(* IEC 61131-3 sources: virtual-bottling-plant/plc/src/generated/bridge, 13 files *)

(* ---- Bridge_Alarms.st ---- *)
(* GENERATED by plc/scripts/gen_plc_io.py from contracts/modbus/plc-io.yaml. Do not edit by hand. *)
(* Alarm table: bit0 active, bit1 acked, bit2 first-out, bits 8-11 prio. *)
PROGRAM Bridge_Alarms
  VAR_EXTERNAL
    G_Alarms : ST_AlarmSummary;
  END_VAR
  VAR
    ALM_T101_BrixOutOfSpec AT %MW601 : INT;
    ALM_T101_CommsLost AT %MW602 : INT;
    ALM_P201_LowTemp AT %MW603 : INT;
    ALM_P201_SteamLow AT %MW604 : INT;
    ALM_P201_CommsLost AT %MW605 : INT;
    ALM_T301_LowLevel AT %MW606 : INT;
    ALM_T301_CommsLost AT %MW607 : INT;
    ALM_F401_NozzleLeak AT %MW608 : INT;
    ALM_F401_CommsLost AT %MW609 : INT;
    ALM_C501_Jam AT %MW610 : INT;
    ALM_C501_Breakdown AT %MW611 : INT;
    ALM_C501_CapsEmpty AT %MW612 : INT;
    ALM_C501_CommsLost AT %MW613 : INT;
    ALM_L601_RollEmpty AT %MW614 : INT;
    ALM_L601_LabelError AT %MW615 : INT;
    ALM_L601_Breakdown AT %MW616 : INT;
    ALM_L601_CommsLost AT %MW617 : INT;
    ALM_Q701_CommsLost AT %MW618 : INT;
    ALM_K801_Jam AT %MW619 : INT;
    ALM_K801_Breakdown AT %MW620 : INT;
    ALM_K801_CommsLost AT %MW621 : INT;
    ALM_LINE_CommsLost AT %MW622 : INT;
  END_VAR
  ALM_T101_BrixOutOfSpec := UINT_TO_INT(G_Alarms.W1);
  ALM_T101_CommsLost := UINT_TO_INT(G_Alarms.W2);
  ALM_P201_LowTemp := UINT_TO_INT(G_Alarms.W3);
  ALM_P201_SteamLow := UINT_TO_INT(G_Alarms.W4);
  ALM_P201_CommsLost := UINT_TO_INT(G_Alarms.W5);
  ALM_T301_LowLevel := UINT_TO_INT(G_Alarms.W6);
  ALM_T301_CommsLost := UINT_TO_INT(G_Alarms.W7);
  ALM_F401_NozzleLeak := UINT_TO_INT(G_Alarms.W8);
  ALM_F401_CommsLost := UINT_TO_INT(G_Alarms.W9);
  ALM_C501_Jam := UINT_TO_INT(G_Alarms.W10);
  ALM_C501_Breakdown := UINT_TO_INT(G_Alarms.W11);
  ALM_C501_CapsEmpty := UINT_TO_INT(G_Alarms.W12);
  ALM_C501_CommsLost := UINT_TO_INT(G_Alarms.W13);
  ALM_L601_RollEmpty := UINT_TO_INT(G_Alarms.W14);
  ALM_L601_LabelError := UINT_TO_INT(G_Alarms.W15);
  ALM_L601_Breakdown := UINT_TO_INT(G_Alarms.W16);
  ALM_L601_CommsLost := UINT_TO_INT(G_Alarms.W17);
  ALM_Q701_CommsLost := UINT_TO_INT(G_Alarms.W18);
  ALM_K801_Jam := UINT_TO_INT(G_Alarms.W19);
  ALM_K801_Breakdown := UINT_TO_INT(G_Alarms.W20);
  ALM_K801_CommsLost := UINT_TO_INT(G_Alarms.W21);
  ALM_LINE_CommsLost := UINT_TO_INT(G_Alarms.W22);
END_PROGRAM

(* ---- Bridge_C501.st ---- *)
(* GENERATED by plc/scripts/gen_plc_io.py from contracts/modbus/plc-io.yaml. Do not edit by hand. *)
(* Status block C501 (%MW200…). *)
PROGRAM Bridge_C501
  VAR_EXTERNAL
    G_In : ST_SimInputs;
    G_Out : ST_SimOutputs;
    G_Status : ST_Status;
    G_Comms : ST_CommsStatus;
    G_Alarms : ST_AlarmSummary;
  END_VAR
  VAR
    C501_State AT %MW200 : INT;
    C501_Mode AT %MW201 : INT;
    C501_StopReason AT %MW202 : INT;
    C501_AlarmWord AT %MW203 : INT;
    C501_CommsOk AT %MW204 : INT;
    C501_Blocked AT %MW205 : INT;
    C501_Starved AT %MW206 : INT;
    C501_Running AT %MW207 : INT;
    C501_Speed AT %MW208 : INT;
    C501_SpeedSP AT %MW209 : INT;
    C501_Torque AT %MW210 : INT;
    C501_LT502_CapHopper AT %MW211 : INT;
  END_VAR
  C501_State := PackMLStateToInt(G_Status.C501.State);
  C501_Mode := PackMLModeToInt(G_Status.C501.Mode);
  C501_StopReason := G_Status.C501.StopReason;
  C501_AlarmWord := G_Alarms.C501_Word;
  C501_CommsOk := BOOL_TO_INT(G_Comms.C501);
  C501_Blocked := BOOL_TO_INT(G_Status.C501.Blocked);
  C501_Starved := BOOL_TO_INT(G_Status.C501.Starved);
  C501_Running := BOOL_TO_INT(G_In.C501_Running);
  C501_Speed := REAL_TO_INT(G_In.C501_Speed);
  C501_SpeedSP := REAL_TO_INT(G_Out.C501_SpeedSP);
  C501_Torque := REAL_TO_INT(G_In.C501_Torque * 100.0);
  C501_LT502_CapHopper := REAL_TO_INT(G_In.LT502_CapHopper * 10.0);
END_PROGRAM

(* ---- Bridge_Commands.st ---- *)
(* GENERATED by plc/scripts/gen_plc_io.py from contracts/modbus/plc-io.yaml. Do not edit by hand. *)
(* One-shot commands: valid in G_Cmd for the scan they arrive, then 0. *)
PROGRAM Bridge_Commands
  VAR_EXTERNAL
    G_Cmd : ST_Commands;
  END_VAR
  VAR
    F401_Cmd AT %MW803 : INT;
    C501_Cmd AT %MW804 : INT;
    L601_Cmd AT %MW805 : INT;
    Q701_Cmd AT %MW806 : INT;
    K801_Cmd AT %MW807 : INT;
    LINE_Cmd AT %MW808 : INT;
    F401_StopReason AT %MW813 : INT;
    C501_StopReason AT %MW814 : INT;
    L601_StopReason AT %MW815 : INT;
    Q701_StopReason AT %MW816 : INT;
    K801_StopReason AT %MW817 : INT;
    AlarmAck AT %MW820 : INT;
    P201_TempSP AT %MW821 : INT;
  END_VAR
  G_Cmd.F401_Cmd := IntToCommand(F401_Cmd);
  F401_Cmd := 0;
  G_Cmd.C501_Cmd := IntToCommand(C501_Cmd);
  C501_Cmd := 0;
  G_Cmd.L601_Cmd := IntToCommand(L601_Cmd);
  L601_Cmd := 0;
  G_Cmd.Q701_Cmd := IntToCommand(Q701_Cmd);
  Q701_Cmd := 0;
  G_Cmd.K801_Cmd := IntToCommand(K801_Cmd);
  K801_Cmd := 0;
  G_Cmd.LINE_Cmd := IntToCommand(LINE_Cmd);
  LINE_Cmd := 0;
  G_Cmd.F401_StopReason := F401_StopReason;
  F401_StopReason := 0;
  G_Cmd.C501_StopReason := C501_StopReason;
  C501_StopReason := 0;
  G_Cmd.L601_StopReason := L601_StopReason;
  L601_StopReason := 0;
  G_Cmd.Q701_StopReason := Q701_StopReason;
  Q701_StopReason := 0;
  G_Cmd.K801_StopReason := K801_StopReason;
  K801_StopReason := 0;
  G_Cmd.AlarmAck := AlarmAck;
  AlarmAck := 0;
  G_Cmd.P201_TempSP := INT_TO_REAL(P201_TempSP) / 10.0;
  P201_TempSP := 0;
END_PROGRAM

(* ---- Bridge_Counters.st ---- *)
(* GENERATED by plc/scripts/gen_plc_io.py from contracts/modbus/plc-io.yaml. Do not edit by hand. *)
(* 32-bit counters (%MD, high word first on Modbus). *)
PROGRAM Bridge_Counters
  VAR_EXTERNAL
    G_In : ST_SimInputs;
    G_Counters : ST_Counters;
  END_VAR
  VAR
    F401_Count AT %MD0 : DINT;
    C501_Count AT %MD1 : DINT;
    L601_Count AT %MD2 : DINT;
    Q701_Count AT %MD3 : DINT;
    Q701_RejectCount AT %MD4 : DINT;
    Q701_GoodCount AT %MD5 : DINT;
    K801_CaseCount AT %MD6 : DINT;
    T101_ConcLotNo AT %MD7 : DINT;
    SIM_TimeMs AT %MD8 : DINT;
  END_VAR
  F401_Count := UDINT_TO_DINT(G_In.F401_Count);
  C501_Count := UDINT_TO_DINT(G_In.C501_Count);
  L601_Count := UDINT_TO_DINT(G_In.L601_Count);
  Q701_Count := UDINT_TO_DINT(G_In.Q701_Count);
  Q701_RejectCount := UDINT_TO_DINT(G_In.Q701_RejectCount);
  Q701_GoodCount := UDINT_TO_DINT(G_Counters.Q701_GoodCount);
  K801_CaseCount := UDINT_TO_DINT(G_In.K801_CaseCount);
  T101_ConcLotNo := UDINT_TO_DINT(G_In.T101_ConcLotNo);
  SIM_TimeMs := UDINT_TO_DINT(G_In.SIM_TimeMs);
END_PROGRAM

(* ---- Bridge_F401.st ---- *)
(* GENERATED by plc/scripts/gen_plc_io.py from contracts/modbus/plc-io.yaml. Do not edit by hand. *)
(* Status block F401 (%MW150…). *)
PROGRAM Bridge_F401
  VAR_EXTERNAL
    G_In : ST_SimInputs;
    G_Out : ST_SimOutputs;
    G_Status : ST_Status;
    G_Comms : ST_CommsStatus;
    G_Alarms : ST_AlarmSummary;
  END_VAR
  VAR
    F401_State AT %MW150 : INT;
    F401_Mode AT %MW151 : INT;
    F401_StopReason AT %MW152 : INT;
    F401_AlarmWord AT %MW153 : INT;
    F401_CommsOk AT %MW154 : INT;
    F401_Blocked AT %MW155 : INT;
    F401_Starved AT %MW156 : INT;
    F401_Running AT %MW157 : INT;
    F401_Speed AT %MW158 : INT;
    F401_SpeedSP AT %MW159 : INT;
    F401_FillTargetG AT %MW160 : INT;
  END_VAR
  F401_State := PackMLStateToInt(G_Status.F401.State);
  F401_Mode := PackMLModeToInt(G_Status.F401.Mode);
  F401_StopReason := G_Status.F401.StopReason;
  F401_AlarmWord := G_Alarms.F401_Word;
  F401_CommsOk := BOOL_TO_INT(G_Comms.F401);
  F401_Blocked := BOOL_TO_INT(G_Status.F401.Blocked);
  F401_Starved := BOOL_TO_INT(G_Status.F401.Starved);
  F401_Running := BOOL_TO_INT(G_In.F401_Running);
  F401_Speed := REAL_TO_INT(G_In.F401_Speed);
  F401_SpeedSP := REAL_TO_INT(G_Out.F401_SpeedSP);
  F401_FillTargetG := REAL_TO_INT(G_Out.F401_FillTargetG * 10.0);
END_PROGRAM

(* ---- Bridge_K801.st ---- *)
(* GENERATED by plc/scripts/gen_plc_io.py from contracts/modbus/plc-io.yaml. Do not edit by hand. *)
(* Status block K801 (%MW350…). *)
PROGRAM Bridge_K801
  VAR_EXTERNAL
    G_In : ST_SimInputs;
    G_Out : ST_SimOutputs;
    G_Status : ST_Status;
    G_Comms : ST_CommsStatus;
    G_Alarms : ST_AlarmSummary;
  END_VAR
  VAR
    K801_State AT %MW350 : INT;
    K801_Mode AT %MW351 : INT;
    K801_StopReason AT %MW352 : INT;
    K801_AlarmWord AT %MW353 : INT;
    K801_CommsOk AT %MW354 : INT;
    K801_Blocked AT %MW355 : INT;
    K801_Starved AT %MW356 : INT;
    K801_Running AT %MW357 : INT;
    K801_Speed AT %MW358 : INT;
    K801_SpeedSP AT %MW359 : INT;
  END_VAR
  K801_State := PackMLStateToInt(G_Status.K801.State);
  K801_Mode := PackMLModeToInt(G_Status.K801.Mode);
  K801_StopReason := G_Status.K801.StopReason;
  K801_AlarmWord := G_Alarms.K801_Word;
  K801_CommsOk := BOOL_TO_INT(G_Comms.K801);
  K801_Blocked := BOOL_TO_INT(G_Status.K801.Blocked);
  K801_Starved := BOOL_TO_INT(G_Status.K801.Starved);
  K801_Running := BOOL_TO_INT(G_In.K801_Running);
  K801_Speed := REAL_TO_INT(G_In.K801_Speed);
  K801_SpeedSP := REAL_TO_INT(G_Out.K801_SpeedSP);
END_PROGRAM

(* ---- Bridge_L601.st ---- *)
(* GENERATED by plc/scripts/gen_plc_io.py from contracts/modbus/plc-io.yaml. Do not edit by hand. *)
(* Status block L601 (%MW250…). *)
PROGRAM Bridge_L601
  VAR_EXTERNAL
    G_In : ST_SimInputs;
    G_Out : ST_SimOutputs;
    G_Status : ST_Status;
    G_Comms : ST_CommsStatus;
    G_Alarms : ST_AlarmSummary;
  END_VAR
  VAR
    L601_State AT %MW250 : INT;
    L601_Mode AT %MW251 : INT;
    L601_StopReason AT %MW252 : INT;
    L601_AlarmWord AT %MW253 : INT;
    L601_CommsOk AT %MW254 : INT;
    L601_Blocked AT %MW255 : INT;
    L601_Starved AT %MW256 : INT;
    L601_Running AT %MW257 : INT;
    L601_Speed AT %MW258 : INT;
    L601_SpeedSP AT %MW259 : INT;
    L601_RollRemaining AT %MW260 : INT;
  END_VAR
  L601_State := PackMLStateToInt(G_Status.L601.State);
  L601_Mode := PackMLModeToInt(G_Status.L601.Mode);
  L601_StopReason := G_Status.L601.StopReason;
  L601_AlarmWord := G_Alarms.L601_Word;
  L601_CommsOk := BOOL_TO_INT(G_Comms.L601);
  L601_Blocked := BOOL_TO_INT(G_Status.L601.Blocked);
  L601_Starved := BOOL_TO_INT(G_Status.L601.Starved);
  L601_Running := BOOL_TO_INT(G_In.L601_Running);
  L601_Speed := REAL_TO_INT(G_In.L601_Speed);
  L601_SpeedSP := REAL_TO_INT(G_Out.L601_SpeedSP);
  L601_RollRemaining := REAL_TO_INT(G_In.L601_RollRemaining);
END_PROGRAM

(* ---- Bridge_LINE.st ---- *)
(* GENERATED by plc/scripts/gen_plc_io.py from contracts/modbus/plc-io.yaml. Do not edit by hand. *)
(* Status block LINE (%MW400…). *)
PROGRAM Bridge_LINE
  VAR_EXTERNAL
    G_In : ST_SimInputs;
    G_Status : ST_Status;
    G_Comms : ST_CommsStatus;
    G_Alarms : ST_AlarmSummary;
  END_VAR
  VAR
    LINE_State AT %MW400 : INT;
    LINE_ActiveAlarmCount AT %MW401 : INT;
    LINE_FirstOutAlarmId AT %MW402 : INT;
    LINE_AlarmWord AT %MW403 : INT;
    LINE_CommsOk AT %MW404 : INT;
    LINE_CV1_Fill AT %MW410 : INT;
    LINE_CV2_Fill AT %MW411 : INT;
    LINE_CV3_Fill AT %MW412 : INT;
    LINE_CV4_Fill AT %MW413 : INT;
    LINE_RecipeId AT %MW420 : INT;
    LINE_RecipeVersion AT %MW421 : INT;
    LINE_ProductCode AT %MW422 : INT;
    LINE_PlcHeartbeat AT %MW449 : INT;
  END_VAR
  LINE_State := PackMLStateToInt(G_Status.LINE.State);
  LINE_ActiveAlarmCount := G_Alarms.ActiveCount;
  LINE_FirstOutAlarmId := G_Alarms.FirstOutId;
  LINE_AlarmWord := G_Alarms.LINE_Word;
  LINE_CommsOk := BOOL_TO_INT(G_Comms.LINE);
  LINE_CV1_Fill := REAL_TO_INT(G_In.CV1_Fill);
  LINE_CV2_Fill := REAL_TO_INT(G_In.CV2_Fill);
  LINE_CV3_Fill := REAL_TO_INT(G_In.CV3_Fill);
  LINE_CV4_Fill := REAL_TO_INT(G_In.CV4_Fill);
  LINE_RecipeId := G_Status.LINE.RecipeId;
  LINE_RecipeVersion := G_Status.LINE.RecipeVersion;
  LINE_ProductCode := G_Status.LINE.ProductCode;
  LINE_PlcHeartbeat := G_Status.LINE.PlcHeartbeat;
END_PROGRAM

(* ---- Bridge_P201.st ---- *)
(* GENERATED by plc/scripts/gen_plc_io.py from contracts/modbus/plc-io.yaml. Do not edit by hand. *)
(* Status block P201 (%MW50…). *)
PROGRAM Bridge_P201
  VAR_EXTERNAL
    G_In : ST_SimInputs;
    G_Out : ST_SimOutputs;
    G_Status : ST_Status;
    G_Comms : ST_CommsStatus;
    G_Alarms : ST_AlarmSummary;
  END_VAR
  VAR
    P201_AlarmWord AT %MW53 : INT;
    P201_CommsOk AT %MW54 : INT;
    P201_TT201_InTemp AT %MW60 : INT;
    P201_TT202_OutTemp AT %MW61 : INT;
    P201_FT201_Flow AT %MW62 : INT;
    P201_PT201_SteamPressure AT %MW63 : INT;
    P201_TCV201_SteamValve AT %MW64 : INT;
    P201_TempSP AT %MW65 : INT;
    P201_XV203_Divert AT %MW66 : INT;
    P201_DivertCount AT %MW67 : INT;
    P201_ForwardFlowOk AT %MW68 : INT;
  END_VAR
  P201_AlarmWord := G_Alarms.P201_Word;
  P201_CommsOk := BOOL_TO_INT(G_Comms.P201);
  P201_TT201_InTemp := REAL_TO_INT(G_In.TT201_InTemp * 10.0);
  P201_TT202_OutTemp := REAL_TO_INT(G_In.TT202_OutTemp * 10.0);
  P201_FT201_Flow := REAL_TO_INT(G_In.FT201_Flow);
  P201_PT201_SteamPressure := REAL_TO_INT(G_In.PT201_SteamPressure * 100.0);
  P201_TCV201_SteamValve := REAL_TO_INT(G_Out.TCV201_SteamValve * 10.0);
  P201_TempSP := REAL_TO_INT(G_Status.P201.TempSP * 10.0);
  P201_XV203_Divert := BOOL_TO_INT(G_Out.XV203_Divert);
  P201_DivertCount := G_Status.P201.DivertCount;
  P201_ForwardFlowOk := BOOL_TO_INT(G_Status.P201.ForwardFlowOk);
END_PROGRAM

(* ---- Bridge_Q701.st ---- *)
(* GENERATED by plc/scripts/gen_plc_io.py from contracts/modbus/plc-io.yaml. Do not edit by hand. *)
(* Status block Q701 (%MW300…). *)
PROGRAM Bridge_Q701
  VAR_EXTERNAL
    G_In : ST_SimInputs;
    G_Out : ST_SimOutputs;
    G_Status : ST_Status;
    G_Comms : ST_CommsStatus;
    G_Alarms : ST_AlarmSummary;
  END_VAR
  VAR
    Q701_State AT %MW300 : INT;
    Q701_Mode AT %MW301 : INT;
    Q701_StopReason AT %MW302 : INT;
    Q701_AlarmWord AT %MW303 : INT;
    Q701_CommsOk AT %MW304 : INT;
    Q701_Blocked AT %MW305 : INT;
    Q701_Starved AT %MW306 : INT;
    Q701_Running AT %MW307 : INT;
    Q701_Speed AT %MW308 : INT;
    Q701_SpeedSP AT %MW309 : INT;
    Q701_RejectLimitG AT %MW310 : INT;
    Q701_WT701_LastWeight AT %MW311 : INT;
    Q701_N01_Seq AT %MW314 : INT;
    Q701_N01_Mean AT %MW315 : INT;
    Q701_N01_Range AT %MW316 : INT;
    Q701_N02_Seq AT %MW317 : INT;
    Q701_N02_Mean AT %MW318 : INT;
    Q701_N02_Range AT %MW319 : INT;
    Q701_N03_Seq AT %MW320 : INT;
    Q701_N03_Mean AT %MW321 : INT;
    Q701_N03_Range AT %MW322 : INT;
    Q701_N04_Seq AT %MW323 : INT;
    Q701_N04_Mean AT %MW324 : INT;
    Q701_N04_Range AT %MW325 : INT;
    Q701_N05_Seq AT %MW326 : INT;
    Q701_N05_Mean AT %MW327 : INT;
    Q701_N05_Range AT %MW328 : INT;
    Q701_N06_Seq AT %MW329 : INT;
    Q701_N06_Mean AT %MW330 : INT;
    Q701_N06_Range AT %MW331 : INT;
    Q701_N07_Seq AT %MW332 : INT;
    Q701_N07_Mean AT %MW333 : INT;
    Q701_N07_Range AT %MW334 : INT;
    Q701_N08_Seq AT %MW335 : INT;
    Q701_N08_Mean AT %MW336 : INT;
    Q701_N08_Range AT %MW337 : INT;
    Q701_N09_Seq AT %MW338 : INT;
    Q701_N09_Mean AT %MW339 : INT;
    Q701_N09_Range AT %MW340 : INT;
    Q701_N10_Seq AT %MW341 : INT;
    Q701_N10_Mean AT %MW342 : INT;
    Q701_N10_Range AT %MW343 : INT;
    Q701_N11_Seq AT %MW344 : INT;
    Q701_N11_Mean AT %MW345 : INT;
    Q701_N11_Range AT %MW346 : INT;
    Q701_N12_Seq AT %MW347 : INT;
    Q701_N12_Mean AT %MW348 : INT;
    Q701_N12_Range AT %MW349 : INT;
  END_VAR
  Q701_State := PackMLStateToInt(G_Status.Q701.State);
  Q701_Mode := PackMLModeToInt(G_Status.Q701.Mode);
  Q701_StopReason := G_Status.Q701.StopReason;
  Q701_AlarmWord := G_Alarms.Q701_Word;
  Q701_CommsOk := BOOL_TO_INT(G_Comms.Q701);
  Q701_Blocked := BOOL_TO_INT(G_Status.Q701.Blocked);
  Q701_Starved := BOOL_TO_INT(G_Status.Q701.Starved);
  Q701_Running := BOOL_TO_INT(G_In.Q701_Running);
  Q701_Speed := REAL_TO_INT(G_In.Q701_Speed);
  Q701_SpeedSP := REAL_TO_INT(G_Out.Q701_SpeedSP);
  Q701_RejectLimitG := REAL_TO_INT(G_Out.Q701_RejectLimitG * 10.0);
  Q701_WT701_LastWeight := REAL_TO_INT(G_In.WT701_LastWeight * 10.0);
  Q701_N01_Seq := UINT_TO_INT(G_In.Q701_N01_Seq);
  Q701_N01_Mean := REAL_TO_INT(G_In.Q701_N01_Mean * 10.0);
  Q701_N01_Range := REAL_TO_INT(G_In.Q701_N01_Range * 10.0);
  Q701_N02_Seq := UINT_TO_INT(G_In.Q701_N02_Seq);
  Q701_N02_Mean := REAL_TO_INT(G_In.Q701_N02_Mean * 10.0);
  Q701_N02_Range := REAL_TO_INT(G_In.Q701_N02_Range * 10.0);
  Q701_N03_Seq := UINT_TO_INT(G_In.Q701_N03_Seq);
  Q701_N03_Mean := REAL_TO_INT(G_In.Q701_N03_Mean * 10.0);
  Q701_N03_Range := REAL_TO_INT(G_In.Q701_N03_Range * 10.0);
  Q701_N04_Seq := UINT_TO_INT(G_In.Q701_N04_Seq);
  Q701_N04_Mean := REAL_TO_INT(G_In.Q701_N04_Mean * 10.0);
  Q701_N04_Range := REAL_TO_INT(G_In.Q701_N04_Range * 10.0);
  Q701_N05_Seq := UINT_TO_INT(G_In.Q701_N05_Seq);
  Q701_N05_Mean := REAL_TO_INT(G_In.Q701_N05_Mean * 10.0);
  Q701_N05_Range := REAL_TO_INT(G_In.Q701_N05_Range * 10.0);
  Q701_N06_Seq := UINT_TO_INT(G_In.Q701_N06_Seq);
  Q701_N06_Mean := REAL_TO_INT(G_In.Q701_N06_Mean * 10.0);
  Q701_N06_Range := REAL_TO_INT(G_In.Q701_N06_Range * 10.0);
  Q701_N07_Seq := UINT_TO_INT(G_In.Q701_N07_Seq);
  Q701_N07_Mean := REAL_TO_INT(G_In.Q701_N07_Mean * 10.0);
  Q701_N07_Range := REAL_TO_INT(G_In.Q701_N07_Range * 10.0);
  Q701_N08_Seq := UINT_TO_INT(G_In.Q701_N08_Seq);
  Q701_N08_Mean := REAL_TO_INT(G_In.Q701_N08_Mean * 10.0);
  Q701_N08_Range := REAL_TO_INT(G_In.Q701_N08_Range * 10.0);
  Q701_N09_Seq := UINT_TO_INT(G_In.Q701_N09_Seq);
  Q701_N09_Mean := REAL_TO_INT(G_In.Q701_N09_Mean * 10.0);
  Q701_N09_Range := REAL_TO_INT(G_In.Q701_N09_Range * 10.0);
  Q701_N10_Seq := UINT_TO_INT(G_In.Q701_N10_Seq);
  Q701_N10_Mean := REAL_TO_INT(G_In.Q701_N10_Mean * 10.0);
  Q701_N10_Range := REAL_TO_INT(G_In.Q701_N10_Range * 10.0);
  Q701_N11_Seq := UINT_TO_INT(G_In.Q701_N11_Seq);
  Q701_N11_Mean := REAL_TO_INT(G_In.Q701_N11_Mean * 10.0);
  Q701_N11_Range := REAL_TO_INT(G_In.Q701_N11_Range * 10.0);
  Q701_N12_Seq := UINT_TO_INT(G_In.Q701_N12_Seq);
  Q701_N12_Mean := REAL_TO_INT(G_In.Q701_N12_Mean * 10.0);
  Q701_N12_Range := REAL_TO_INT(G_In.Q701_N12_Range * 10.0);
END_PROGRAM

(* ---- Bridge_Recipe.st ---- *)
(* GENERATED by plc/scripts/gen_plc_io.py from contracts/modbus/plc-io.yaml. Do not edit by hand. *)
(* Recipe download block and Req/Ack/Nak handshake (contracts.md §2). *)
PROGRAM Bridge_Recipe
  VAR_EXTERNAL
    G_RecipeReq : ST_RecipeRequest;
    G_RecipeResp : ST_RecipeResponse;
  END_VAR
  VAR
    Recipe_Req AT %MW900 : INT;
    RecipeId AT %MW903 : INT;
    RecipeVersion AT %MW904 : INT;
    ProductCode AT %MW905 : INT;
    BrixTarget AT %MW906 : INT;
    BrixTol AT %MW907 : INT;
    ConcRatio AT %MW908 : INT;
    FillTargetG AT %MW909 : INT;
    LineSpeed AT %MW910 : INT;
    CapTorque AT %MW911 : INT;
    Recipe_Ack AT %MW901 : INT;
    Recipe_Nak AT %MW902 : INT;
  END_VAR
  G_RecipeReq.Recipe_Req := Recipe_Req <> 0;
  G_RecipeReq.RecipeId := RecipeId;
  G_RecipeReq.RecipeVersion := RecipeVersion;
  G_RecipeReq.ProductCode := ProductCode;
  G_RecipeReq.BrixTarget := INT_TO_REAL(BrixTarget) / 100.0;
  G_RecipeReq.BrixTol := INT_TO_REAL(BrixTol) / 100.0;
  G_RecipeReq.ConcRatio := INT_TO_REAL(ConcRatio) / 1000.0;
  G_RecipeReq.FillTargetG := INT_TO_REAL(FillTargetG) / 10.0;
  G_RecipeReq.LineSpeed := LineSpeed;
  G_RecipeReq.CapTorque := INT_TO_REAL(CapTorque) / 100.0;
  Recipe_Ack := BOOL_TO_INT(G_RecipeResp.Recipe_Ack);
  Recipe_Nak := RecipeNakToInt(G_RecipeResp.Recipe_Nak);
END_PROGRAM

(* ---- Bridge_T101.st ---- *)
(* GENERATED by plc/scripts/gen_plc_io.py from contracts/modbus/plc-io.yaml. Do not edit by hand. *)
(* Status block T101 (%MW0…). *)
PROGRAM Bridge_T101
  VAR_EXTERNAL
    G_In : ST_SimInputs;
    G_Out : ST_SimOutputs;
    G_Status : ST_Status;
    G_Comms : ST_CommsStatus;
    G_Alarms : ST_AlarmSummary;
  END_VAR
  VAR
    T101_Phase AT %MW0 : INT;
    T101_AlarmWord AT %MW3 : INT;
    T101_CommsOk AT %MW4 : INT;
    T101_LT101_Level AT %MW10 : INT;
    T101_AT101_Brix AT %MW11 : INT;
    T101_BatchNo AT %MW12 : INT;
    T101_ProductCode AT %MW13 : INT;
    T101_BatchBrix AT %MW14 : INT;
    T101_BrixOk AT %MW15 : INT;
    T101_BatchActive AT %MW16 : INT;
    T101_M101_Agitator AT %MW17 : INT;
  END_VAR
  T101_Phase := BatchPhaseToInt(G_Status.T101.Phase);
  T101_AlarmWord := G_Alarms.T101_Word;
  T101_CommsOk := BOOL_TO_INT(G_Comms.T101);
  T101_LT101_Level := REAL_TO_INT(G_In.LT101_Level * 10.0);
  T101_AT101_Brix := REAL_TO_INT(G_In.AT101_Brix * 100.0);
  T101_BatchNo := G_Status.T101.BatchNo;
  T101_ProductCode := G_Status.T101.ProductCode;
  T101_BatchBrix := REAL_TO_INT(G_Status.T101.BatchBrix * 100.0);
  T101_BrixOk := BOOL_TO_INT(G_Status.T101.BrixOk);
  T101_BatchActive := BOOL_TO_INT(G_Status.T101.BatchActive);
  T101_M101_Agitator := BOOL_TO_INT(G_Out.M101_Agitator);
END_PROGRAM

(* ---- Bridge_T301.st ---- *)
(* GENERATED by plc/scripts/gen_plc_io.py from contracts/modbus/plc-io.yaml. Do not edit by hand. *)
(* Status block T301 (%MW100…). *)
PROGRAM Bridge_T301
  VAR_EXTERNAL
    G_In : ST_SimInputs;
    G_Status : ST_Status;
    G_Comms : ST_CommsStatus;
    G_Alarms : ST_AlarmSummary;
  END_VAR
  VAR
    T301_AlarmWord AT %MW103 : INT;
    T301_CommsOk AT %MW104 : INT;
    T301_LT301_Level AT %MW110 : INT;
    T301_FillerPermissive AT %MW111 : INT;
  END_VAR
  T301_AlarmWord := G_Alarms.T301_Word;
  T301_CommsOk := BOOL_TO_INT(G_Comms.T301);
  T301_LT301_Level := REAL_TO_INT(G_In.LT301_Level * 10.0);
  T301_FillerPermissive := BOOL_TO_INT(G_Status.T301.FillerPermissive);
END_PROGRAM
